Fanuc KAREL source: KT00796.KL

PROGRAM KT00796
%NOLOCKGROUP
VAR
  I1: INTEGER
  I2: INTEGER
  OUT: INTEGER
BEGIN
  I1 = 2
  I2 = 3
  I1 = 2
  I2 = 3
  OUT = EXP(I1)
END KT00796
